Fanuc TP program (LS listing): NamePr.LS

/PROG  NamePr
/ATTR
OWNER		= MNEDITOR;
COMMENT		= "RoboDK sequence";
PROG_SIZE	= 0;
CREATE		= DATE 31-12-14  TIME 12:00:00;
MODIFIED	= DATE 31-12-14  TIME 12:00:00;
FILE_NAME	= NamePr;
VERSION		= 0;
LINE_COUNT	= 23;
MEMORY_SIZE	= 0;
PROTECT		= READ_WRITE;
TCD:  STACK_SIZE	= 0,
      TASK_PRIORITY	= 50,
      TIME_SLICE	= 0,
      BUSY_LAMP_OFF	= 0,
      ABORT_REQUEST	= 0,
      PAUSE_REQUEST	= 0;
DEFAULT_GROUP	= 1,*,*,*,*;
CONTROL_CODE	= 00000000 00000000;
/MN
   1:  ! Program generated by RoboDK v6.0.7 for Fanuc ARC Mate 100iD/8 ;
   2:  ! L on XX/XX/XXXX 18:00:00 ;
   3:  ! Using nominal kinematics. ;
   4:  PR[9,1]=1234.570 ;
   5:  PR[9,2]=-98.765 ;
   6:  PR[9,3]=50.500 ;
   7:  PR[9,4]=0.000 ;
   8:  PR[9,5]=0.000 ;
   9:  PR[9,6]=30.000 ;
  10:  UFRAME[9]=PR[9] ;
  11:  UFRAME_NUM=9 ;
  12:  PR[9,1]=10.000 ;
  13:  PR[9,2]=20.000 ;
  14:  PR[9,3]=150.000 ;
  15:  PR[9,4]=0.000 ;
  16:  PR[9,5]=0.000 ;
  17:  PR[9,6]=0.000 ;
  18:  UTOOL[9]=PR[9] ;
  19:  UTOOL_NUM=9 ;
  20:J P[1] 20% FINE ;
  21:L P[2] 200mm/sec FINE ;
  22:C P[3]
       P[4] 200mm/sec FINE ;
  23:J P[5] 20% FINE ;
/POS
P[1]{
   GP1:
    UF : 9, UT : 9,
	J1=    0.000 deg,	J2=    -10.000 deg,	J3=    20.000 deg,
	J4=    0.000 deg,	J5=    30.000 deg,	J6=    0.000 deg
};
P[2]{
   GP1:
    UF : 9, UT : 9,        CONFIG : 'N U T, 0, 0, 0',
	X =  -607.850  mm,	Y =   543.849  mm,	Z =   363.215  mm,
	W =  -165.000 deg,	P =    50.000 deg,	R =   150.000 deg
};
P[3]{
   GP1:
    UF : 9, UT : 9,        CONFIG : 'N U T, 0, 0, 0',
	X =  -602.951  mm,	Y =   596.788  mm,	Z =   316.595  mm,
	W =  -165.000 deg,	P =    50.000 deg,	R =   150.000 deg
};
P[4]{
   GP1:
    UF : 9, UT : 9,        CONFIG : 'N U T, 0, 0, 0',
	X =  -663.517  mm,	Y =   575.988  mm,	Z =   286.611  mm,
	W =  -165.000 deg,	P =    50.000 deg,	R =   150.000 deg
};
P[5]{
   GP1:
    UF : 9, UT : 9,
	J1=    20.000 deg,	J2=    -10.000 deg,	J3=    20.000 deg,
	J4=    0.000 deg,	J5=    30.000 deg,	J6=    0.000 deg
};
/END
